TEXTLIST TextList_RecipeRootFolder
  0 = 'PLC'
  1 = 'Develop 1'
  2 = 'Develop 2'
  3 = 'Develop 3'
  4 = 'Develop 4'
   = ''
END_TEXTLIST

(* stored: Version 1.1.0.1, ProductVersion 3.1.4024.12
   TextList TextList_RecipeRootFolder: Id {040425d0-1796-4d18-8fae-b52d0c6d3c57} *)
